Fanuc KAREL source: kt00366.KL

-- PROVISIONAL review KL for V940-1; original PC SHA256 93b5e3a8137715b037a881379a6dda2fd15c1deb816ab41fcf58e6cb462ad226
-- Incomplete behavior may be omitted. Consult companion uncertainty JSON. Do not deploy.
PROGRAM KT00366
%NOLOCKGROUP
VAR
  I1 : INTEGER
  R2 : REAL
  OUT : BOOLEAN
BEGIN
  -- V9_ZERO_TABLE_METADATA_HINT layout=0001; no indexed target words; source/name/runtime held
  -- UNRESOLVED_PC offsets 5-16; opcodes 2E,23
  -- UNRESOLVED_PC offsets 21-32; opcodes 2E,23
  -- UNRESOLVED_PC offsets 37-59; opcodes 21,21,29,64,29,70,23
  -- UNRESOLVED_PC offsets 64-68; opcodes 7F
END KT00366
